(* IEC 61131-3 sources: SortJet_MasterSPS_Aufbau.fbsproj/Device.device.xml.v3^/Plc Logic.plclogic.xml.v3^/Application.application.xml.v3^/05_Sicherheitstechnik, 2 files *)

(* ---- Interface_SLC.prg.st ---- *)
(* METADATA
{
	"v3Meta": {
		"objectGuid": "ccad9978-fd7c-48d9-8d85-dc1a7581631d"
	}
}
*)
PROGRAM Interface_SLC

VAR_INPUT

  // BOOL
  bpResetOperatorAcknowledge : BOOL;
  bpEDMFehlerAktiv           : BOOL;

END_VAR

VAR_OUTPUT

  // BOOL
  bpOperatorAcknowledgeRequested : BOOL; // HINWEIS: Mindestens ein Safety IO Modul hat einen Fehler, es ist erforderlich das der Anwender wissendlich diesen Zustand zuruecksetzt

END_VAR

VAR

  // BOOLEAN
  bpVisuResetEDM                  : BOOL := FALSE;
  bpVisuResetFSoEMaster           : BOOL;
  bpVisuResetNothalt              : BOOL;
  bResetDurchSK                   : BOOL;
  ablSKAbgefallen                 : ARRAY[1..16] OF BOOL;

  // WORD
  wIndex                         : WORD := 0;
  wlbitPos                       : WORD;

  // TIMER
  toflResetOA                                    : TOF;
  toflSKQuittiert                                : ARRAY[cERSTER_SICHERHEITSKREIS..cLETZTER_SICHERHEITSKREIS] OF tof;
  tonlSKKomplettAbgefallen                       : ARRAY[cERSTER_SICHERHEITSKREIS..cLETZTER_SICHERHEITSKREIS] OF TON;

  // TRIGGER
  rtlMeldungQuittierungDurchBedienerErforderlich : R_TRIG;
  rtlResetOA                                     : R_TRIG;
  rtlSKQuittiert                                 : ARRAY[cERSTER_SICHERHEITSKREIS..cLETZTER_SICHERHEITSKREIS] OF R_TRIG;;

END_VAR

//-------------------------------------------------------------------------------------------------
// AKTIONEN
//-------------------------------------------------------------------------------------------------
OperatorAcknowledge();
SK_Hilfsvariablen();
Meldungen();
ToSLC();
ToPLC();
END_PROGRAM

(* ---- NotHalt.prg.st ---- *)
(* METADATA
{
	"v3Meta": {
		"objectGuid": "69a82f5e-5606-42e6-b3a3-559b5ec715fe"
	}
}
*)
PROGRAM NotHalt
VAR_INPUT

  // BOOL
  bpEingangNotHaltOK        : BOOL; // Not-Halt ok von SLC

  // WORD
  wMeldungsnummer           : WORD;

END_VAR
VAR_OUTPUT

  // BOOLE
  bpNotHaltOK               : BOOL;
  bpTasterNothaltQuittieren : BOOL;

END_VAR
VAR

  // BOOL
  blResetNotHalt     : BOOL := FALSE;

  // RS-FLIP FLOP
  NotHaltAusgeloest : SR;
  NotHaltQuittieren : RS;

  // TIMER
  tonlNotHaltAusgeloest : TON;

END_VAR
VAR
  // HARDWARE EINGAENGE
  in_bTasterNothaltQuittieren             AT %I* : BOOL; // Taster zum Quittieren des Nothalts und Reset der Safety-Module

  // HARDWARE AUSGAENGE
  out_bLeuchtdruckTasterNotHaltAusgeloest  AT %Q* : BOOL;

END_VAR
VAR CONSTANT

  // TIME VALUE
  cZEIT_NOTAUS_VERZOEGERUNG : TIME := T#100MS;

END_VAR
//-------------------------------------------------------------------------------------------------
// Taster
//-------------------------------------------------------------------------------------------------

// Leuchtdruck Taster am CAB
out_bLeuchtdruckTasterNotHaltAusgeloest := NOT bpNotHaltOK OR ( Interface_SLC.bpEDMFehlerAktiv AND gbFlashbit05sec );
bpTasterNothaltQuittieren := in_bTasterNothaltQuittieren OR Interface_SLC.bpVisuResetNothalt;

//-------------------------------------------------------------------------------------------------
// BAUSTEIN: AKTIONEN
//-------------------------------------------------------------------------------------------------
Meldungen();

//-------------------------------------------------------------------------------------------------
// BAUSTEIN: LOGIK
//-------------------------------------------------------------------------------------------------
// Kurze Verzoegerung das alle Signale durchgeschaltet haben
tonlNotHaltAusgeloest( IN := ( NOT bpEingangNotHaltOK OR bgSicherheitstechnikBruecken ),
                       PT := cZEIT_NOTAUS_VERZOEGERUNG );

// NotHalt OK bilden
bpNotHaltOK := (   NOT NotHaltAusgeloest.Q1
                 OR Visu_Notaus_OK
                 OR bgSicherheitstechnikBruecken );

(* Hinweis:
   - Merker das der Notaus ausgeloest wurde
     => Bistabiele Funktion in der das  "set" dominant ist
*)
NotHaltAusgeloest( SET1 := tonlNotHaltAusgeloest.Q,
                   RESET:= blResetNotHalt );

(* Hinweis:
   - Merker das der Taster "Quittierung Notaus" betaetigt wurde
     => Bistabiele Funktion in der das  "reset" dominant ist
*)
NotHaltQuittieren( SET   := ( in_bTasterNothaltQuittieren OR Interface_SLC.bpVisuResetNothalt ) ,
                   RESET1:= NOT NotHaltAusgeloest.Q1);

IF ( NotHaltQuittieren.Q1
     AND NOT tonlNotHaltAusgeloest.Q )
THEN
  blResetNotHalt := TRUE;
ELSE
  blResetNotHalt := FALSE;
END_IF
END_PROGRAM
